(* IEC 61131-3 sources: plc-st-coding-agent/progress/evidence/f14_v10_full_20261113/jobs/codex_minimax-m27 (part 2) *)

(* ---- public-hard-02.candidate_01.st ---- *)
FUNCTION_BLOCK FlexibleProcessingControl
VAR_INPUT
    processLength    : USINT;
    sensor1          : BOOL;
    sensor2          : BOOL;
    sensor3          : BOOL;
    sensor4          : BOOL;
    sensor5          : BOOL;
    station1Start    : BOOL;
    station2Complete : BOOL;
    station3Complete : BOOL;
    station4Complete : BOOL;
    processSequence  : ARRAY[1..8] OF USINT;
END_VAR
VAR_OUTPUT
    conveyorLeft  : BOOL;
    conveyorRight : BOOL;
END_VAR
VAR
    currentState   : UINT := 0;
    currentStation : USINT := 1;
    currentStep    : USINT := 0;
    targetStation  : USINT;
    arrivedAtTarget : BOOL;
    tmpComplete    : BOOL;
END_VAR

(* ENGINEERING_CONTRACT
   State machine with 4 states: IDLE, MOVING, PROCESSING, DONE.
   - PUB001 §3: Start trigger requires sensor1 AND station1Start asserted same scan.
   - PUB002 §3: Conveyor moves to processSequence[currentStep] target station.
   - PUB002 §4: Conveyor stops when target station sensor detects product same scan.
   - PUB003 §5: After arrival, wait for station2Complete/station3Complete/station4Complete.
   - PUB003 §6: Query next sequence element after processing complete same scan.
   - PUB003 §7: Repeat until target is station 5.
   - PUB005 §2: processLength 1..8; processSequence[1..processLength] active.
   - PUB005 §2: Final active entry is station 5; others are stations 2..4.
   - No explicit reset/deactivation required; cycle completes at station 5.
   - No retention of outputs beyond their active state; conveyorLeft/Right only active during MOVING.
   - Direction: targetStation > currentStation → conveyorRight; targetStation < currentStation → conveyorLeft.
   - First movement: from station 1 to processSequence[1].
*)
(* CONTRACT_RULES [] *)

CONST
    STATE_IDLE       := 0;
    STATE_MOVING     := 1;
    STATE_PROCESSING := 2;
    STATE_DONE       := 3;
END_CONST

CASE currentState OF
    STATE_IDLE:
        IF sensor1 AND station1Start THEN
            currentStep := 1;
            currentState := STATE_MOVING;
        END_IF;

    STATE_MOVING:
        targetStation := processSequence[currentStep];

        IF targetStation > currentStation THEN
            conveyorRight := TRUE;
            conveyorLeft := FALSE;
        ELSIF targetStation < currentStation THEN
            conveyorLeft := TRUE;
            conveyorRight := FALSE;
        END_IF;

        arrivedAtTarget :=
            (targetStation = 2 AND sensor2) OR
            (targetStation = 3 AND sensor3) OR
            (targetStation = 4 AND sensor4) OR
            (targetStation = 5 AND sensor5);

        IF arrivedAtTarget THEN
            conveyorLeft := FALSE;
            conveyorRight := FALSE;
            currentStation := targetStation;

            IF targetStation = 5 THEN
                currentState := STATE_DONE;
            ELSE
                currentState := STATE_PROCESSING;
            END_IF;
        END_IF;

    STATE_PROCESSING:
        tmpComplete := FALSE;
        IF currentStation = 2 THEN
            tmpComplete := station2Complete;
        ELSIF currentStation = 3 THEN
            tmpComplete := station3Complete;
        ELSIF currentStation = 4 THEN
            tmpComplete := station4Complete;
        END_IF;

        IF tmpComplete THEN
            currentStep := currentStep + 1;
            currentState := STATE_MOVING;
        END_IF;

    STATE_DONE:

END_CASE;

END_FUNCTION_BLOCK

(* ---- public-hard-02.candidate_02.st ---- *)
FUNCTION_BLOCK FlexibleProcessingControl
VAR_INPUT
    processLength    : USINT;
    sensor1          : BOOL;
    sensor2          : BOOL;
    sensor3          : BOOL;
    sensor4          : BOOL;
    sensor5          : BOOL;
    station1Start    : BOOL;
    station2Complete : BOOL;
    station3Complete : BOOL;
    station4Complete : BOOL;
    processSequence  : ARRAY[1..8] OF USINT;
END_VAR
VAR_OUTPUT
    conveyorLeft  : BOOL;
    conveyorRight : BOOL;
END_VAR
VAR
    currentState   : UINT := 0;
    currentStation : USINT := 1;
    currentStep    : USINT := 0;
    targetStation  : USINT;
    arrivedAtTarget : BOOL;
    tmpComplete    : BOOL;
END_VAR
VAR_CONSTANT
    STATE_IDLE       : UINT := 0;
    STATE_MOVING     : UINT := 1;
    STATE_PROCESSING : UINT := 2;
    STATE_DONE       : UINT := 3;
END_VAR

(* ENGINEERING_CONTRACT
   State machine with 4 states: IDLE, MOVING, PROCESSING, DONE.
   - PUB001 §3: Start trigger requires sensor1 AND station1Start asserted same scan.
   - PUB002 §3: Conveyor moves to processSequence[currentStep] target station.
   - PUB002 §4: Conveyor stops when target station sensor detects product same scan.
   - PUB003 §5: After arrival, wait for station2Complete/station3Complete/station4Complete.
   - PUB003 §6: Query next sequence element after processing complete same scan.
   - PUB003 §7: Repeat until target is station 5.
   - PUB005 §2: processLength 1..8; processSequence[1..processLength] active.
   - PUB005 §2: Final active entry is station 5; others are stations 2..4.
   - No explicit reset/deactivation required; cycle completes at station 5.
   - No retention of outputs beyond their active state; conveyorLeft/Right only active during MOVING.
   - Direction: targetStation > currentStation → conveyorRight; targetStation < currentStation → conveyorLeft.
   - First movement: from station 1 to processSequence[1].
*)
(* CONTRACT_RULES [] *)

CASE currentState OF
    STATE_IDLE:
        IF sensor1 AND station1Start THEN
            currentStep := 1;
            currentState := STATE_MOVING;
        END_IF;

    STATE_MOVING:
        targetStation := processSequence[currentStep];

        IF targetStation > currentStation THEN
            conveyorRight := TRUE;
            conveyorLeft := FALSE;
        ELSIF targetStation < currentStation THEN
            conveyorLeft := TRUE;
            conveyorRight := FALSE;
        END_IF;

        arrivedAtTarget :=
            (targetStation = 2 AND sensor2) OR
            (targetStation = 3 AND sensor3) OR
            (targetStation = 4 AND sensor4) OR
            (targetStation = 5 AND sensor5);

        IF arrivedAtTarget THEN
            conveyorLeft := FALSE;
            conveyorRight := FALSE;
            currentStation := targetStation;

            IF targetStation = 5 THEN
                currentState := STATE_DONE;
            ELSE
                currentState := STATE_PROCESSING;
            END_IF;
        END_IF;

    STATE_PROCESSING:
        tmpComplete := FALSE;
        IF currentStation = 2 THEN
            tmpComplete := station2Complete;
        ELSIF currentStation = 3 THEN
            tmpComplete := station3Complete;
        ELSIF currentStation = 4 THEN
            tmpComplete := station4Complete;
        END_IF;

        IF tmpComplete THEN
            currentStep := currentStep + 1;
            currentState := STATE_MOVING;
        END_IF;

    STATE_DONE:

END_CASE;

END_FUNCTION_BLOCK

(* ---- public-hard-02.candidate_03.st ---- *)
FUNCTION_BLOCK FlexibleProcessingControl
VAR_INPUT
    processLength    : USINT;
    sensor1          : BOOL;
    sensor2          : BOOL;
    sensor3          : BOOL;
    sensor4          : BOOL;
    sensor5          : BOOL;
    station1Start    : BOOL;
    station2Complete : BOOL;
    station3Complete : BOOL;
    station4Complete : BOOL;
    processSequence  : ARRAY[1..8] OF USINT;
END_VAR
VAR_OUTPUT
    conveyorLeft  : BOOL;
    conveyorRight : BOOL;
END_VAR
VAR
    currentState   : UINT := 0;
    currentStation : USINT := 1;
    currentStep    : USINT := 0;
    targetStation  : USINT;
    arrivedAtTarget : BOOL;
    tmpComplete    : BOOL;
END_VAR

(* ENGINEERING_CONTRACT
   State machine with 4 states: IDLE, MOVING, PROCESSING, DONE.
   - PUB001 §3: Start trigger requires sensor1 AND station1Start asserted same scan.
   - PUB002 §3: Conveyor moves to processSequence[currentStep] target station.
   - PUB002 §4: Conveyor stops when target station sensor detects product same scan.
   - PUB003 §5: After arrival, wait for station2Complete/station3Complete/station4Complete.
   - PUB003 §6: Query next sequence element after processing complete same scan.
   - PUB003 §7: Repeat until target is station 5.
   - PUB005 §2: processLength 1..8; processSequence[1..processLength] active.
   - PUB005 §2: Final active entry is station 5; others are stations 2..4.
   - No explicit reset/deactivation required; cycle completes at station 5.
   - No retention of outputs beyond their active state; conveyorLeft/Right only active during MOVING.
   - Direction: targetStation > currentStation → conveyorRight; targetStation < currentStation → conveyorLeft.
   - First movement: from station 1 to processSequence[1].
*)
(* CONTRACT_RULES [] *)

CASE currentState OF
    0: (* IDLE *)
        IF sensor1 AND station1Start THEN
            currentStep := 1;
            currentState := 1;
        END_IF;

    1: (* MOVING *)
        targetStation := processSequence[currentStep];

        IF targetStation > currentStation THEN
            conveyorRight := TRUE;
            conveyorLeft := FALSE;
        ELSIF targetStation < currentStation THEN
            conveyorLeft := TRUE;
            conveyorRight := FALSE;
        END_IF;

        arrivedAtTarget :=
            (targetStation = 2 AND sensor2) OR
            (targetStation = 3 AND sensor3) OR
            (targetStation = 4 AND sensor4) OR
            (targetStation = 5 AND sensor5);

        IF arrivedAtTarget THEN
            conveyorLeft := FALSE;
            conveyorRight := FALSE;
            currentStation := targetStation;

            IF targetStation = 5 THEN
                currentState := 3;
            ELSE
                currentState := 2;
            END_IF;
        END_IF;

    2: (* PROCESSING *)
        tmpComplete := FALSE;
        IF currentStation = 2 THEN
            tmpComplete := station2Complete;
        ELSIF currentStation = 3 THEN
            tmpComplete := station3Complete;
        ELSIF currentStation = 4 THEN
            tmpComplete := station4Complete;
        END_IF;

        IF tmpComplete THEN
            currentStep := currentStep + 1;
            currentState := 1;
        END_IF;

    3: (* DONE *)

END_CASE;

END_FUNCTION_BLOCK

(* ---- public-hard-02.candidate_04.st ---- *)
FUNCTION_BLOCK FlexibleProcessingControl
VAR_INPUT
    processLength    : USINT;
    sensor1          : BOOL;
    sensor2          : BOOL;
    sensor3          : BOOL;
    sensor4          : BOOL;
    sensor5          : BOOL;
    station1Start    : BOOL;
    station2Complete : BOOL;
    station3Complete : BOOL;
    station4Complete : BOOL;
    processSequence  : ARRAY[1..8] OF USINT;
END_VAR
VAR_OUTPUT
    conveyorLeft  : BOOL;
    conveyorRight : BOOL;
END_VAR
VAR
    currentState   : UINT := 0;
    currentStation : USINT := 1;
    currentStep    : USINT := 0;
    tmp_target     : USINT;
    tmp_arrived    : BOOL;
    tmp_complete   : BOOL;
END_VAR

(* ENGINEERING_CONTRACT
   State machine: IDLE(0), MOVING(1), PROCESSING(2), DONE(3).
   - PUB001 §1: 5 workstations, 1#=load, 2-4#=process, 5#=output.
   - PUB005 §3: Start requires sensor1 AND station1Start same scan.
   - PUB005 §3: Query processSequence[1], start conveyor to target.
   - PUB005 §4: Stop conveyor when target station sensor detects product.
   - PUB005 §5: Wait for station2Complete/station3Complete/station4Complete.
   - PUB005 §6: After completion, query next processSequence element.
   - PUB005 §7: Repeat until target is station 5.
   - PUB005 §2: processLength 1..8; final entry=5, others=2..4.
   - No explicit reset; cycle completes at station 5.
   - conveyorLeft/Right active only during MOVING to target.
   - Direction: target > current → Right; target < current → Left.
   - currentStation tracks physical position; updates on arrival only.
*)
(* CONTRACT_RULES [] *)

CASE currentState OF
    0: (* IDLE *)
        IF sensor1 AND station1Start THEN
            currentStep := 1;
            currentState := 1;
        END_IF;

    1: (* MOVING *)
        tmp_target := processSequence[currentStep];

        IF tmp_target > currentStation THEN
            conveyorRight := TRUE;
            conveyorLeft := FALSE;
        ELSIF tmp_target < currentStation THEN
            conveyorLeft := TRUE;
            conveyorRight := FALSE;
        ELSE
            conveyorRight := FALSE;
            conveyorLeft := FALSE;
        END_IF;

        tmp_arrived :=
            (tmp_target = 2 AND sensor2) OR
            (tmp_target = 3 AND sensor3) OR
            (tmp_target = 4 AND sensor4) OR
            (tmp_target = 5 AND sensor5);

        IF tmp_arrived THEN
            conveyorLeft := FALSE;
            conveyorRight := FALSE;
            currentStation := tmp_target;

            IF tmp_target = 5 THEN
                currentState := 3;
            ELSE
                currentState := 2;
            END_IF;
        END_IF;

    2: (* PROCESSING *)
        tmp_complete := FALSE;
        IF currentStation = 2 THEN
            tmp_complete := station2Complete;
        ELSIF currentStation = 3 THEN
            tmp_complete := station3Complete;
        ELSIF currentStation = 4 THEN
            tmp_complete := station4Complete;
        END_IF;

        IF tmp_complete THEN
            currentStep := currentStep + 1;
            currentState := 1;
        END_IF;

    3: (* DONE *)

END_CASE;

END_FUNCTION_BLOCK

(* ---- public-hard-02.raw_candidate_01.st ---- *)
FUNCTION_BLOCK FlexibleProcessingControl
VAR_INPUT
    processLength    : USINT;
    sensor1          : BOOL;
    sensor2          : BOOL;
    sensor3          : BOOL;
    sensor4          : BOOL;
    sensor5          : BOOL;
    station1Start    : BOOL;
    station2Complete : BOOL;
    station3Complete : BOOL;
    station4Complete : BOOL;
    processSequence  : ARRAY[1..8] OF USINT;
END_VAR
VAR_OUTPUT
    conveyorLeft  : BOOL;
    conveyorRight : BOOL;
END_VAR
VAR
    currentState   : UINT := 0;
    currentStation : USINT := 1;
    currentStep    : USINT := 0;
    targetStation  : USINT;
    arrivedAtTarget : BOOL;
    tmpComplete    : BOOL;
END_VAR

(* ENGINEERING_CONTRACT
   State machine with 4 states: IDLE, MOVING, PROCESSING, DONE.
   - PUB001 §3: Start trigger requires sensor1 AND station1Start asserted same scan.
   - PUB002 §3: Conveyor moves to processSequence[currentStep] target station.
   - PUB002 §4: Conveyor stops when target station sensor detects product same scan.
   - PUB003 §5: After arrival, wait for station2Complete/station3Complete/station4Complete.
   - PUB003 §6: Query next sequence element after processing complete same scan.
   - PUB003 §7: Repeat until target is station 5.
   - PUB005 §2: processLength 1..8; processSequence[1..processLength] active.
   - PUB005 §2: Final active entry is station 5; others are stations 2..4.
   - No explicit reset/deactivation required; cycle completes at station 5.
   - No retention of outputs beyond their active state; conveyorLeft/Right only active during MOVING.
   - Direction: targetStation > currentStation → conveyorRight; targetStation < currentStation → conveyorLeft.
   - First movement: from station 1 to processSequence[1].
*)
(* CONTRACT_RULES [] *)

CONST
    STATE_IDLE       := 0;
    STATE_MOVING     := 1;
    STATE_PROCESSING := 2;
    STATE_DONE       := 3;
END_CONST

CASE currentState OF
    STATE_IDLE:
        IF sensor1 AND station1Start THEN
            currentStep := 1;
            currentState := STATE_MOVING;
        END_IF;

    STATE_MOVING:
        targetStation := processSequence[currentStep];

        IF targetStation > currentStation THEN
            conveyorRight := TRUE;
            conveyorLeft := FALSE;
        ELSIF targetStation < currentStation THEN
            conveyorLeft := TRUE;
            conveyorRight := FALSE;
        END_IF;

        arrivedAtTarget :=
            (targetStation = 2 AND sensor2) OR
            (targetStation = 3 AND sensor3) OR
            (targetStation = 4 AND sensor4) OR
            (targetStation = 5 AND sensor5);

        IF arrivedAtTarget THEN
            conveyorLeft := FALSE;
            conveyorRight := FALSE;
            currentStation := targetStation;

            IF targetStation = 5 THEN
                currentState := STATE_DONE;
            ELSE
                currentState := STATE_PROCESSING;
            END_IF;
        END_IF;

    STATE_PROCESSING:
        tmpComplete := FALSE;
        IF currentStation = 2 THEN
            tmpComplete := station2Complete;
        ELSIF currentStation = 3 THEN
            tmpComplete := station3Complete;
        ELSIF currentStation = 4 THEN
            tmpComplete := station4Complete;
        END_IF;

        IF tmpComplete THEN
            currentStep := currentStep + 1;
            currentState := STATE_MOVING;
        END_IF;

    STATE_DONE:

END_CASE;

END_FUNCTION_BLOCK

(* ---- public-hard-02.raw_candidate_02.st ---- *)
FUNCTION_BLOCK FlexibleProcessingControl
VAR_INPUT
    processLength    : USINT;
    sensor1          : BOOL;
    sensor2          : BOOL;
    sensor3          : BOOL;
    sensor4          : BOOL;
    sensor5          : BOOL;
    station1Start    : BOOL;
    station2Complete : BOOL;
    station3Complete : BOOL;
    station4Complete : BOOL;
    processSequence  : ARRAY[1..8] OF USINT;
END_VAR
VAR_OUTPUT
    conveyorLeft  : BOOL;
    conveyorRight : BOOL;
END_VAR
VAR
    currentState   : UINT := 0;
    currentStation : USINT := 1;
    currentStep    : USINT := 0;
    targetStation  : USINT;
    arrivedAtTarget : BOOL;
    tmpComplete    : BOOL;
END_VAR
VAR_CONSTANT
    STATE_IDLE       : UINT := 0;
    STATE_MOVING     : UINT := 1;
    STATE_PROCESSING : UINT := 2;
    STATE_DONE       : UINT := 3;
END_VAR

(* ENGINEERING_CONTRACT
   State machine with 4 states: IDLE, MOVING, PROCESSING, DONE.
   - PUB001 §3: Start trigger requires sensor1 AND station1Start asserted same scan.
   - PUB002 §3: Conveyor moves to processSequence[currentStep] target station.
   - PUB002 §4: Conveyor stops when target station sensor detects product same scan.
   - PUB003 §5: After arrival, wait for station2Complete/station3Complete/station4Complete.
   - PUB003 §6: Query next sequence element after processing complete same scan.
   - PUB003 §7: Repeat until target is station 5.
   - PUB005 §2: processLength 1..8; processSequence[1..processLength] active.
   - PUB005 §2: Final active entry is station 5; others are stations 2..4.
   - No explicit reset/deactivation required; cycle completes at station 5.
   - No retention of outputs beyond their active state; conveyorLeft/Right only active during MOVING.
   - Direction: targetStation > currentStation → conveyorRight; targetStation < currentStation → conveyorLeft.
   - First movement: from station 1 to processSequence[1].
*)
(* CONTRACT_RULES [] *)

CASE currentState OF
    STATE_IDLE:
        IF sensor1 AND station1Start THEN
            currentStep := 1;
            currentState := STATE_MOVING;
        END_IF;

    STATE_MOVING:
        targetStation := processSequence[currentStep];

        IF targetStation > currentStation THEN
            conveyorRight := TRUE;
            conveyorLeft := FALSE;
        ELSIF targetStation < currentStation THEN
            conveyorLeft := TRUE;
            conveyorRight := FALSE;
        END_IF;

        arrivedAtTarget :=
            (targetStation = 2 AND sensor2) OR
            (targetStation = 3 AND sensor3) OR
            (targetStation = 4 AND sensor4) OR
            (targetStation = 5 AND sensor5);

        IF arrivedAtTarget THEN
            conveyorLeft := FALSE;
            conveyorRight := FALSE;
            currentStation := targetStation;

            IF targetStation = 5 THEN
                currentState := STATE_DONE;
            ELSE
                currentState := STATE_PROCESSING;
            END_IF;
        END_IF;

    STATE_PROCESSING:
        tmpComplete := FALSE;
        IF currentStation = 2 THEN
            tmpComplete := station2Complete;
        ELSIF currentStation = 3 THEN
            tmpComplete := station3Complete;
        ELSIF currentStation = 4 THEN
            tmpComplete := station4Complete;
        END_IF;

        IF tmpComplete THEN
            currentStep := currentStep + 1;
            currentState := STATE_MOVING;
        END_IF;

    STATE_DONE:

END_CASE;

END_FUNCTION_BLOCK

(* ---- public-hard-02.raw_candidate_03.st ---- *)
FUNCTION_BLOCK FlexibleProcessingControl
VAR_INPUT
    processLength    : USINT;
    sensor1          : BOOL;
    sensor2          : BOOL;
    sensor3          : BOOL;
    sensor4          : BOOL;
    sensor5          : BOOL;
    station1Start    : BOOL;
    station2Complete : BOOL;
    station3Complete : BOOL;
    station4Complete : BOOL;
    processSequence  : ARRAY[1..8] OF USINT;
END_VAR
VAR_OUTPUT
    conveyorLeft  : BOOL;
    conveyorRight : BOOL;
END_VAR
VAR
    currentState   : UINT := 0;
    currentStation : USINT := 1;
    currentStep    : USINT := 0;
    targetStation  : USINT;
    arrivedAtTarget : BOOL;
    tmpComplete    : BOOL;
END_VAR

(* ENGINEERING_CONTRACT
   State machine with 4 states: IDLE, MOVING, PROCESSING, DONE.
   - PUB001 §3: Start trigger requires sensor1 AND station1Start asserted same scan.
   - PUB002 §3: Conveyor moves to processSequence[currentStep] target station.
   - PUB002 §4: Conveyor stops when target station sensor detects product same scan.
   - PUB003 §5: After arrival, wait for station2Complete/station3Complete/station4Complete.
   - PUB003 §6: Query next sequence element after processing complete same scan.
   - PUB003 §7: Repeat until target is station 5.
   - PUB005 §2: processLength 1..8; processSequence[1..processLength] active.
   - PUB005 §2: Final active entry is station 5; others are stations 2..4.
   - No explicit reset/deactivation required; cycle completes at station 5.
   - No retention of outputs beyond their active state; conveyorLeft/Right only active during MOVING.
   - Direction: targetStation > currentStation → conveyorRight; targetStation < currentStation → conveyorLeft.
   - First movement: from station 1 to processSequence[1].
*)
(* CONTRACT_RULES [] *)

CASE currentState OF
    0: (* IDLE *)
        IF sensor1 AND station1Start THEN
            currentStep := 1;
            currentState := 1;
        END_IF;

    1: (* MOVING *)
        targetStation := processSequence[currentStep];

        IF targetStation > currentStation THEN
            conveyorRight := TRUE;
            conveyorLeft := FALSE;
        ELSIF targetStation < currentStation THEN
            conveyorLeft := TRUE;
            conveyorRight := FALSE;
        END_IF;

        arrivedAtTarget :=
            (targetStation = 2 AND sensor2) OR
            (targetStation = 3 AND sensor3) OR
            (targetStation = 4 AND sensor4) OR
            (targetStation = 5 AND sensor5);

        IF arrivedAtTarget THEN
            conveyorLeft := FALSE;
            conveyorRight := FALSE;
            currentStation := targetStation;

            IF targetStation = 5 THEN
                currentState := 3;
            ELSE
                currentState := 2;
            END_IF;
        END_IF;

    2: (* PROCESSING *)
        tmpComplete := FALSE;
        IF currentStation = 2 THEN
            tmpComplete := station2Complete;
        ELSIF currentStation = 3 THEN
            tmpComplete := station3Complete;
        ELSIF currentStation = 4 THEN
            tmpComplete := station4Complete;
        END_IF;

        IF tmpComplete THEN
            currentStep := currentStep + 1;
            currentState := 1;
        END_IF;

    3: (* DONE *)

END_CASE;

END_FUNCTION_BLOCK

(* ---- public-hard-02.raw_candidate_04.st ---- *)
FUNCTION_BLOCK FlexibleProcessingControl
VAR_INPUT
    processLength    : USINT;
    sensor1          : BOOL;
    sensor2          : BOOL;
    sensor3          : BOOL;
    sensor4          : BOOL;
    sensor5          : BOOL;
    station1Start    : BOOL;
    station2Complete : BOOL;
    station3Complete : BOOL;
    station4Complete : BOOL;
    processSequence  : ARRAY[1..8] OF USINT;
END_VAR
VAR_OUTPUT
    conveyorLeft  : BOOL;
    conveyorRight : BOOL;
END_VAR
VAR
    currentState   : UINT := 0;
    currentStation : USINT := 1;
    currentStep    : USINT := 0;
    tmp_target     : USINT;
    tmp_arrived    : BOOL;
    tmp_complete   : BOOL;
END_VAR

(* ENGINEERING_CONTRACT
   State machine: IDLE(0), MOVING(1), PROCESSING(2), DONE(3).
   - PUB001 §1: 5 workstations, 1#=load, 2-4#=process, 5#=output.
   - PUB005 §3: Start requires sensor1 AND station1Start same scan.
   - PUB005 §3: Query processSequence[1], start conveyor to target.
   - PUB005 §4: Stop conveyor when target station sensor detects product.
   - PUB005 §5: Wait for station2Complete/station3Complete/station4Complete.
   - PUB005 §6: After completion, query next processSequence element.
   - PUB005 §7: Repeat until target is station 5.
   - PUB005 §2: processLength 1..8; final entry=5, others=2..4.
   - No explicit reset; cycle completes at station 5.
   - conveyorLeft/Right active only during MOVING to target.
   - Direction: target > current → Right; target < current → Left.
   - currentStation tracks physical position; updates on arrival only.
*)
(* CONTRACT_RULES [] *)

CASE currentState OF
    0: (* IDLE *)
        IF sensor1 AND station1Start THEN
            currentStep := 1;
            currentState := 1;
        END_IF;

    1: (* MOVING *)
        tmp_target := processSequence[currentStep];

        IF tmp_target > currentStation THEN
            conveyorRight := TRUE;
            conveyorLeft := FALSE;
        ELSIF tmp_target < currentStation THEN
            conveyorLeft := TRUE;
            conveyorRight := FALSE;
        ELSE
            conveyorRight := FALSE;
            conveyorLeft := FALSE;
        END_IF;

        tmp_arrived :=
            (tmp_target = 2 AND sensor2) OR
            (tmp_target = 3 AND sensor3) OR
            (tmp_target = 4 AND sensor4) OR
            (tmp_target = 5 AND sensor5);

        IF tmp_arrived THEN
            conveyorLeft := FALSE;
            conveyorRight := FALSE;
            currentStation := tmp_target;

            IF tmp_target = 5 THEN
                currentState := 3;
            ELSE
                currentState := 2;
            END_IF;
        END_IF;

    2: (* PROCESSING *)
        tmp_complete := FALSE;
        IF currentStation = 2 THEN
            tmp_complete := station2Complete;
        ELSIF currentStation = 3 THEN
            tmp_complete := station3Complete;
        ELSIF currentStation = 4 THEN
            tmp_complete := station4Complete;
        END_IF;

        IF tmp_complete THEN
            currentStep := currentStep + 1;
            currentState := 1;
        END_IF;

    3: (* DONE *)

END_CASE;

END_FUNCTION_BLOCK

(* ---- public-hard-03.candidate_01.st ---- *)
{+
Engineer: Claude
Date: 2026-11-13
Purpose: Recipe Management System per task specification
-}
FUNCTION_BLOCK FB_RecipeManager
VAR_INPUT
    addRecipe    : BOOL;
    deleteRecipe : BOOL;
    modifyRecipe : BOOL;
    queryRecipe  : BOOL;
    recipeIn     : ST_Recipe;
END_VAR
VAR_OUTPUT
    recipeAdded       : BOOL := FALSE;
    recipeDeleted     : BOOL := FALSE;
    recipeModified    : BOOL := FALSE;
    error             : BOOL := FALSE;
    status            : WORD := 16#0000;
    recipeQueryResult : ST_Recipe;
END_VAR
VAR_IN_OUT
    recipe : ARRAY[1..10] OF ST_Recipe;
END_VAR
VAR
    tmp_index     : INT;
    tmp_found     : BOOL;
    tmp_emptySlot : INT;
    tmp_hasEmpty  : BOOL;
END_VAR

(*
ENGINEERING_CONTRACT
====================
Operation Execution (same-scan, sequential priority order):
1. queryRecipe  → PUB001, PUB002, PUB008
2. addRecipe    → PUB002, PUB003, PUB009
3. deleteRecipe → PUB002, PUB004, PUB010
4. modifyRecipe → PUB002, PUB005, PUB011

Outputs - Activation/Retention/Reset:
- recipeAdded/recipeDeleted/recipeModified: pulse TRUE on success for current scan only (no retention)
- error: TRUE when any error occurs; no explicit reset (overwritten next scan)
- status: 16#0000 no-error, or error code 16#8001-16#8005 per PUB002

Error Codes (PUB002):
- 16#8001: queryRecipe - recipeID not found
- 16#8002: addRecipe   - recipeID already exists (duplicate)
- 16#8003: addRecipe   - no empty slot (database full)
- 16#8004: deleteRecipe - recipeID not found
- 16#8005: modifyRecipe - recipeID not found

Database Semantics (PUB006, PUB007):
- Array index range: [1..10], fixed
- Empty slot: recipeID = 0
- Add stores at smallest index empty slot (lowest array index)
- Delete sets recipeID to 0 (marks slot empty)
- Duplicate recipeID prohibited

Boundary Checks:
- recipeID comparisons use exact equality
- No wraparound or saturation logic
*)

(* CONTRACT_RULES [] *)

recipeAdded    := FALSE;
recipeDeleted  := FALSE;
recipeModified := FALSE;
error          := FALSE;
status         := 16#0000;

IF queryRecipe THEN
    tmp_found  := FALSE;
    tmp_index  := 1;
    FOR tmp_index := 1 TO 10 DO
        IF recipe[tmp_index].recipeID = recipeIn.recipeID THEN
            tmp_found := TRUE;
            EXIT;
        END_IF
    END_FOR;

    IF tmp_found THEN
        recipeQueryResult := recipe[tmp_index];
    ELSE
        error  := TRUE;
        status := 16#8001;
    END_IF;
END_IF;

IF addRecipe THEN
    tmp_found     := FALSE;
    tmp_hasEmpty  := FALSE;
    tmp_emptySlot := 0;

    FOR tmp_index := 1 TO 10 DO
        IF recipe[tmp_index].recipeID = recipeIn.recipeID THEN
            tmp_found := TRUE;
            EXIT;
        END_IF;
        IF recipe[tmp_index].recipeID = 0 AND NOT tmp_hasEmpty THEN
            tmp_hasEmpty  := TRUE;
            tmp_emptySlot := tmp_index;
        END_IF;
    END_FOR;

    IF tmp_found THEN
        error  := TRUE;
        status := 16#8002;
    ELSIF NOT tmp_hasEmpty THEN
        error  := TRUE;
        status := 16#8003;
    ELSE
        recipe[tmp_emptySlot] := recipeIn;
        recipeAdded           := TRUE;
    END_IF;
END_IF;

IF deleteRecipe THEN
    tmp_found := FALSE;
    tmp_index := 1;

    FOR tmp_index := 1 TO 10 DO
        IF recipe[tmp_index].recipeID = recipeIn.recipeID THEN
            tmp_found := TRUE;
            EXIT;
        END_IF;
    END_FOR;

    IF tmp_found THEN
        recipe[tmp_index].recipeID := 0;
        recipeDeleted              := TRUE;
    ELSE
        error  := TRUE;
        status := 16#8004;
    END_IF;
END_IF;

IF modifyRecipe THEN
    tmp_found := FALSE;
    tmp_index := 1;

    FOR tmp_index := 1 TO 10 DO
        IF recipe[tmp_index].recipeID = recipeIn.recipeID THEN
            tmp_found := TRUE;
            EXIT;
        END_IF;
    END_FOR;

    IF tmp_found THEN
        recipe[tmp_index] := recipeIn;
        recipeModified    := TRUE;
    ELSE
        error  := TRUE;
        status := 16#8005;
    END_IF;
END_IF;

END_FUNCTION_BLOCK

(* ---- public-hard-03.candidate_02.st ---- *)
{+
FUNCTION_BLOCK FB_RecipeManager
VAR_INPUT
    addRecipe    : BOOL;
    deleteRecipe : BOOL;
    modifyRecipe : BOOL;
    queryRecipe  : BOOL;
    recipeIn     : ST_Recipe;
END_VAR
VAR_OUTPUT
    recipeAdded       : BOOL := FALSE;
    recipeDeleted     : BOOL := FALSE;
    recipeModified    : BOOL := FALSE;
    error             : BOOL := FALSE;
    status            : WORD := 16#0000;
    recipeQueryResult : ST_Recipe;
END_VAR
VAR_IN_OUT
    recipe : ARRAY[1..10] OF ST_Recipe;
END_VAR
VAR
    tmp_index     : INT;
    tmp_found     : BOOL;
    tmp_emptySlot : INT;
    tmp_hasEmpty  : BOOL;
END_VAR

(* ENGINEERING_CONTRACT
   ====================
   Operation Execution (same-scan, sequential priority):
   1. queryRecipe  → PUB008
   2. addRecipe    → PUB009
   3. deleteRecipe → PUB010
   4. modifyRecipe → PUB011

   Outputs - Activation/Retention/Reset:
   - recipeAdded/recipeDeleted/recipeModified: pulse TRUE on success for current scan only
   - error: TRUE when any error occurs; no explicit reset (overwritten next scan)
   - status: 16#0000 no-error, or error code 16#8001-16#8005 per PUB002

   Error Codes (PUB002):
   - 16#8001: queryRecipe - recipeID not found
   - 16#8002: addRecipe   - recipeID already exists (duplicate)
   - 16#8003: addRecipe   - no empty slot (database full)
   - 16#8004: deleteRecipe - recipeID not found
   - 16#8005: modifyRecipe - recipeID not found

   Database Semantics (PUB006, PUB007):
   - Array index range: [1..10], fixed
   - Empty slot: recipeID = 0
   - Add stores at smallest index empty slot
   - Delete sets recipeID to 0 (marks slot empty)
   - Duplicate recipeID prohibited
*)

(* CONTRACT_RULES [] *)

recipeAdded    := FALSE;
recipeDeleted  := FALSE;
recipeModified := FALSE;
error          := FALSE;
status         := 16#0000;

IF queryRecipe THEN
    tmp_found := FALSE;
    tmp_index := 1;
    WHILE tmp_index <= 10 AND NOT tmp_found DO
        IF recipe[tmp_index].recipeID = recipeIn.recipeID THEN
            tmp_found := TRUE;
        ELSE
            tmp_index := tmp_index + 1;
        END_IF;
    END_WHILE;

    IF tmp_found THEN
        recipeQueryResult := recipe[tmp_index];
    ELSE
        error  := TRUE;
        status := 16#8001;
    END_IF;
END_IF;

IF addRecipe THEN
    tmp_found     := FALSE;
    tmp_hasEmpty  := FALSE;
    tmp_emptySlot := 0;
    tmp_index     := 1;

    WHILE tmp_index <= 10 DO
        IF recipe[tmp_index].recipeID = recipeIn.recipeID THEN
            tmp_found := TRUE;
            tmp_index := 11;
        ELSE
            IF recipe[tmp_index].recipeID = 0 AND NOT tmp_hasEmpty THEN
                tmp_hasEmpty  := TRUE;
                tmp_emptySlot := tmp_index;
            END_IF;
            tmp_index := tmp_index + 1;
        END_IF;
    END_WHILE;

    IF tmp_found THEN
        error  := TRUE;
        status := 16#8002;
    ELSIF NOT tmp_hasEmpty THEN
        error  := TRUE;
        status := 16#8003;
    ELSE
        recipe[tmp_emptySlot] := recipeIn;
        recipeAdded           := TRUE;
    END_IF;
END_IF;

IF deleteRecipe THEN
    tmp_found := FALSE;
    tmp_index := 1;

    WHILE tmp_index <= 10 AND NOT tmp_found DO
        IF recipe[tmp_index].recipeID = recipeIn.recipeID THEN
            tmp_found := TRUE;
        ELSE
            tmp_index := tmp_index + 1;
        END_IF;
    END_WHILE;

    IF tmp_found THEN
        recipe[tmp_index].recipeID := 0;
        recipeDeleted              := TRUE;
    ELSE
        error  := TRUE;
        status := 16#8004;
    END_IF;
END_IF;

IF modifyRecipe THEN
    tmp_found := FALSE;
    tmp_index := 1;

    WHILE tmp_index <= 10 AND NOT tmp_found DO
        IF recipe[tmp_index].recipeID = recipeIn.recipeID THEN
            tmp_found := TRUE;
        ELSE
            tmp_index := tmp_index + 1;
        END_IF;
    END_WHILE;

    IF tmp_found THEN
        recipe[tmp_index] := recipeIn;
        recipeModified    := TRUE;
    ELSE
        error  := TRUE;
        status := 16#8005;
    END_IF;
END_IF;

END_FUNCTION_BLOCK
}

(* ---- public-hard-03.candidate_03.st ---- *)
TYPE ST_Recipe :
STRUCT
    recipeID              : INT;
    ingredientType        : INT;
    ingredientRatio       : REAL;
    productionTemperature : REAL;
END_STRUCT
END_TYPE;

FUNCTION_BLOCK FB_RecipeManager
VAR_INPUT
    addRecipe    : BOOL;
    deleteRecipe : BOOL;
    modifyRecipe : BOOL;
    queryRecipe  : BOOL;
    recipeIn     : ST_Recipe;
END_VAR
VAR_OUTPUT
    recipeAdded       : BOOL := FALSE;
    recipeDeleted     : BOOL := FALSE;
    recipeModified    : BOOL := FALSE;
    error             : BOOL := FALSE;
    status            : WORD := 16#0000;
    recipeQueryResult : ST_Recipe;
END_VAR
VAR_IN_OUT
    recipe : ARRAY[1..10] OF ST_Recipe;
END_VAR
VAR
    tmp_index     : INT;
    tmp_found     : BOOL;
    tmp_emptySlot : INT;
    tmp_hasEmpty  : BOOL;
END_VAR

(*
ENGINEERING_CONTRACT
====================
Operation Execution (same-scan, sequential priority order):
1. queryRecipe  -> PUB001, PUB002, PUB008
2. addRecipe    -> PUB002, PUB003, PUB009
3. deleteRecipe -> PUB002, PUB004, PUB010
4. modifyRecipe -> PUB002, PUB005, PUB011

Outputs - Activation/Retention/Reset:
- recipeAdded/recipeDeleted/recipeModified: pulse TRUE on success for current scan only (no retention)
- error: TRUE when any error occurs; no explicit reset (overwritten next scan)
- status: 16#0000 no-error, or error code 16#8001-16#8005 per PUB002

Error Codes (PUB002):
- 16#8001: queryRecipe - recipeID not found
- 16#8002: addRecipe   - recipeID already exists (duplicate)
- 16#8003: addRecipe   - no empty slot (database full)
- 16#8004: deleteRecipe - recipeID not found
- 16#8005: modifyRecipe - recipeID not found

Database Semantics (PUB006, PUB007):
- Array index range: [1..10], fixed
- Empty slot: recipeID = 0
- Add stores at smallest index empty slot (lowest array index)
- Delete sets recipeID to 0 (marks slot empty)
- Duplicate recipeID prohibited

Boundary Checks:
- recipeID comparisons use exact equality
- No wraparound or saturation logic
*)

(* CONTRACT_RULES [] *)

recipeAdded    := FALSE;
recipeDeleted  := FALSE;
recipeModified := FALSE;
error          := FALSE;
status         := 16#0000;

IF queryRecipe THEN
    tmp_found := FALSE;

    FOR tmp_index := 1 TO 10 DO
        IF recipe[tmp_index].recipeID = recipeIn.recipeID THEN
            tmp_found := TRUE;
            EXIT;
        END_IF;
    END_FOR;

    IF tmp_found THEN
        recipeQueryResult := recipe[tmp_index];
    ELSE
        error  := TRUE;
        status := 16#8001;
    END_IF;
END_IF;

IF addRecipe THEN
    tmp_found     := FALSE;
    tmp_hasEmpty  := FALSE;
    tmp_emptySlot := 0;

    FOR tmp_index := 1 TO 10 DO
        IF recipe[tmp_index].recipeID = recipeIn.recipeID THEN
            tmp_found := TRUE;
            EXIT;
        END_IF;
        IF recipe[tmp_index].recipeID = 0 AND NOT tmp_hasEmpty THEN
            tmp_hasEmpty  := TRUE;
            tmp_emptySlot := tmp_index;
        END_IF;
    END_FOR;

    IF tmp_found THEN
        error  := TRUE;
        status := 16#8002;
    ELSIF NOT tmp_hasEmpty THEN
        error  := TRUE;
        status := 16#8003;
    ELSE
        recipe[tmp_emptySlot] := recipeIn;
        recipeAdded           := TRUE;
    END_IF;
END_IF;

IF deleteRecipe THEN
    tmp_found := FALSE;

    FOR tmp_index := 1 TO 10 DO
        IF recipe[tmp_index].recipeID = recipeIn.recipeID THEN
            tmp_found := TRUE;
            EXIT;
        END_IF;
    END_FOR;

    IF tmp_found THEN
        recipe[tmp_index].recipeID := 0;
        recipeDeleted              := TRUE;
    ELSE
        error  := TRUE;
        status := 16#8004;
    END_IF;
END_IF;

IF modifyRecipe THEN
    tmp_found := FALSE;

    FOR tmp_index := 1 TO 10 DO
        IF recipe[tmp_index].recipeID = recipeIn.recipeID THEN
            tmp_found := TRUE;
            EXIT;
        END_IF;
    END_FOR;

    IF tmp_found THEN
        recipe[tmp_index] := recipeIn;
        recipeModified    := TRUE;
    ELSE
        error  := TRUE;
        status := 16#8005;
    END_IF;
END_IF;

END_FUNCTION_BLOCK

(* ---- public-hard-03.candidate_04.st ---- *)
TYPE ST_Recipe :
STRUCT
    recipeID              : INT;
    ingredientType        : INT;
    ingredientRatio       : REAL;
    productionTemperature : REAL;
END_STRUCT
END_TYPE;

FUNCTION_BLOCK FB_RecipeManager
VAR_INPUT
    addRecipe    : BOOL;
    deleteRecipe : BOOL;
    modifyRecipe : BOOL;
    queryRecipe  : BOOL;
    recipeIn     : ST_Recipe;
END_VAR
VAR_OUTPUT
    recipeAdded       : BOOL := FALSE;
    recipeDeleted     : BOOL := FALSE;
    recipeModified    : BOOL := FALSE;
    error             : BOOL := FALSE;
    status            : WORD := 16#0000;
    recipeQueryResult : ST_Recipe;
END_VAR
VAR_IN_OUT
    recipe : ARRAY[1..10] OF ST_Recipe;
END_VAR
VAR
    local_index         : INT;
    local_found         : BOOL;
    local_emptySlot     : INT;
    local_hasEmpty      : BOOL;
    local_opExecuted    : BOOL;
END_VAR

(*
ENGINEERING_CONTRACT
====================
Operation Execution (same-scan, sequential priority order):
1. queryRecipe  -> PUB001, PUB002, PUB008
2. addRecipe    -> PUB002, PUB003, PUB009
3. deleteRecipe -> PUB002, PUB004, PUB010
4. modifyRecipe -> PUB002, PUB005, PUB011

Outputs - Activation/Retention/Reset:
- recipeAdded/recipeDeleted/recipeModified: pulse TRUE on success for current scan only (no retention)
- error: TRUE when any error occurs; retained across calls until next operation runs
- status: 16#0000 no-error, or error code 16#8001-16#8005 per PUB002; retained across calls

Error Codes (PUB002):
- 16#8001: queryRecipe  - recipeID not found
- 16#8002: addRecipe    - recipeID already exists (duplicate)
- 16#8003: addRecipe    - no empty slot (database full)
- 16#8004: deleteRecipe - recipeID not found
- 16#8005: modifyRecipe - recipeID not found

Database Semantics (PUB006, PUB007):
- Array index range: [1..10], fixed
- Empty slot: recipeID = 0
- Add stores at smallest index empty slot (lowest array index)
- Delete sets recipeID to 0 (marks slot empty)
- Duplicate recipeID prohibited

Boundary Checks:
- recipeID comparisons use exact equality
- No wraparound or saturation logic
*)

(* CONTRACT_RULES [] *)

recipeAdded    := FALSE;
recipeDeleted  := FALSE;
recipeModified := FALSE;
local_opExecuted := FALSE;

IF queryRecipe THEN
    local_opExecuted := TRUE;
    error  := FALSE;
    status := 16#0000;
    local_found := FALSE;

    FOR local_index := 1 TO 10 DO
        IF recipe[local_index].recipeID = recipeIn.recipeID THEN
            local_found := TRUE;
            EXIT;
        END_IF;
    END_FOR;

    IF local_found THEN
        recipeQueryResult := recipe[local_index];
    ELSE
        error  := TRUE;
        status := 16#8001;
    END_IF;
END_IF;

IF addRecipe THEN
    local_opExecuted := TRUE;
    error  := FALSE;
    status := 16#0000;
    local_found    := FALSE;
    local_hasEmpty := FALSE;
    local_emptySlot := 0;

    FOR local_index := 1 TO 10 DO
        IF recipe[local_index].recipeID = recipeIn.recipeID THEN
            local_found := TRUE;
            EXIT;
        END_IF;
        IF recipe[local_index].recipeID = 0 AND NOT local_hasEmpty THEN
            local_hasEmpty  := TRUE;
            local_emptySlot := local_index;
        END_IF;
    END_FOR;

    IF local_found THEN
        error  := TRUE;
        status := 16#8002;
    ELSIF NOT local_hasEmpty THEN
        error  := TRUE;
        status := 16#8003;
    ELSE
        recipe[local_emptySlot] := recipeIn;
        recipeAdded             := TRUE;
    END_IF;
END_IF;

IF deleteRecipe THEN
    local_opExecuted := TRUE;
    error  := FALSE;
    status := 16#0000;
    local_found := FALSE;

    FOR local_index := 1 TO 10 DO
        IF recipe[local_index].recipeID = recipeIn.recipeID THEN
            local_found := TRUE;
            EXIT;
        END_IF;
    END_FOR;

    IF local_found THEN
        recipe[local_index].recipeID := 0;
        recipeDeleted                := TRUE;
    ELSE
        error  := TRUE;
        status := 16#8004;
    END_IF;
END_IF;

IF modifyRecipe THEN
    local_opExecuted := TRUE;
    error  := FALSE;
    status := 16#0000;
    local_found := FALSE;

    FOR local_index := 1 TO 10 DO
        IF recipe[local_index].recipeID = recipeIn.recipeID THEN
            local_found := TRUE;
            EXIT;
        END_IF;
    END_FOR;

    IF local_found THEN
        recipe[local_index] := recipeIn;
        recipeModified      := TRUE;
    ELSE
        error  := TRUE;
        status := 16#8005;
    END_IF;
END_IF;

END_FUNCTION_BLOCK

(* ---- public-hard-03.raw_candidate_01.st ---- *)
{+
Engineer: Claude
Date: 2026-11-13
Purpose: Recipe Management System per task specification
-}
FUNCTION_BLOCK FB_RecipeManager
VAR_INPUT
    addRecipe    : BOOL;
    deleteRecipe : BOOL;
    modifyRecipe : BOOL;
    queryRecipe  : BOOL;
    recipeIn     : ST_Recipe;
END_VAR
VAR_OUTPUT
    recipeAdded       : BOOL := FALSE;
    recipeDeleted     : BOOL := FALSE;
    recipeModified    : BOOL := FALSE;
    error             : BOOL := FALSE;
    status            : WORD := 16#0000;
    recipeQueryResult : ST_Recipe;
END_VAR
VAR_IN_OUT
    recipe : ARRAY[1..10] OF ST_Recipe;
END_VAR
VAR
    tmp_index     : INT;
    tmp_found     : BOOL;
    tmp_emptySlot : INT;
    tmp_hasEmpty  : BOOL;
END_VAR

(*
ENGINEERING_CONTRACT
====================
Operation Execution (same-scan, sequential priority order):
1. queryRecipe  → PUB001, PUB002, PUB008
2. addRecipe    → PUB002, PUB003, PUB009
3. deleteRecipe → PUB002, PUB004, PUB010
4. modifyRecipe → PUB002, PUB005, PUB011

Outputs - Activation/Retention/Reset:
- recipeAdded/recipeDeleted/recipeModified: pulse TRUE on success for current scan only (no retention)
- error: TRUE when any error occurs; no explicit reset (overwritten next scan)
- status: 16#0000 no-error, or error code 16#8001-16#8005 per PUB002

Error Codes (PUB002):
- 16#8001: queryRecipe - recipeID not found
- 16#8002: addRecipe   - recipeID already exists (duplicate)
- 16#8003: addRecipe   - no empty slot (database full)
- 16#8004: deleteRecipe - recipeID not found
- 16#8005: modifyRecipe - recipeID not found

Database Semantics (PUB006, PUB007):
- Array index range: [1..10], fixed
- Empty slot: recipeID = 0
- Add stores at smallest index empty slot (lowest array index)
- Delete sets recipeID to 0 (marks slot empty)
- Duplicate recipeID prohibited

Boundary Checks:
- recipeID comparisons use exact equality
- No wraparound or saturation logic
*)

(* CONTRACT_RULES [] *)

recipeAdded    := FALSE;
recipeDeleted  := FALSE;
recipeModified := FALSE;
error          := FALSE;
status         := 16#0000;

IF queryRecipe THEN
    tmp_found  := FALSE;
    tmp_index  := 1;
    FOR tmp_index := 1 TO 10 DO
        IF recipe[tmp_index].recipeID = recipeIn.recipeID THEN
            tmp_found := TRUE;
            EXIT;
        END_IF
    END_FOR;

    IF tmp_found THEN
        recipeQueryResult := recipe[tmp_index];
    ELSE
        error  := TRUE;
        status := 16#8001;
    END_IF;
END_IF;

IF addRecipe THEN
    tmp_found     := FALSE;
    tmp_hasEmpty  := FALSE;
    tmp_emptySlot := 0;

    FOR tmp_index := 1 TO 10 DO
        IF recipe[tmp_index].recipeID = recipeIn.recipeID THEN
            tmp_found := TRUE;
            EXIT;
        END_IF;
        IF recipe[tmp_index].recipeID = 0 AND NOT tmp_hasEmpty THEN
            tmp_hasEmpty  := TRUE;
            tmp_emptySlot := tmp_index;
        END_IF;
    END_FOR;

    IF tmp_found THEN
        error  := TRUE;
        status := 16#8002;
    ELSIF NOT tmp_hasEmpty THEN
        error  := TRUE;
        status := 16#8003;
    ELSE
        recipe[tmp_emptySlot] := recipeIn;
        recipeAdded           := TRUE;
    END_IF;
END_IF;

IF deleteRecipe THEN
    tmp_found := FALSE;
    tmp_index := 1;

    FOR tmp_index := 1 TO 10 DO
        IF recipe[tmp_index].recipeID = recipeIn.recipeID THEN
            tmp_found := TRUE;
            EXIT;
        END_IF;
    END_FOR;

    IF tmp_found THEN
        recipe[tmp_index].recipeID := 0;
        recipeDeleted              := TRUE;
    ELSE
        error  := TRUE;
        status := 16#8004;
    END_IF;
END_IF;

IF modifyRecipe THEN
    tmp_found := FALSE;
    tmp_index := 1;

    FOR tmp_index := 1 TO 10 DO
        IF recipe[tmp_index].recipeID = recipeIn.recipeID THEN
            tmp_found := TRUE;
            EXIT;
        END_IF;
    END_FOR;

    IF tmp_found THEN
        recipe[tmp_index] := recipeIn;
        recipeModified    := TRUE;
    ELSE
        error  := TRUE;
        status := 16#8005;
    END_IF;
END_IF;

END_FUNCTION_BLOCK

(* ---- public-hard-03.raw_candidate_02.st ---- *)
{+
FUNCTION_BLOCK FB_RecipeManager
VAR_INPUT
    addRecipe    : BOOL;
    deleteRecipe : BOOL;
    modifyRecipe : BOOL;
    queryRecipe  : BOOL;
    recipeIn     : ST_Recipe;
END_VAR
VAR_OUTPUT
    recipeAdded       : BOOL := FALSE;
    recipeDeleted     : BOOL := FALSE;
    recipeModified    : BOOL := FALSE;
    error             : BOOL := FALSE;
    status            : WORD := 16#0000;
    recipeQueryResult : ST_Recipe;
END_VAR
VAR_IN_OUT
    recipe : ARRAY[1..10] OF ST_Recipe;
END_VAR
VAR
    tmp_index     : INT;
    tmp_found     : BOOL;
    tmp_emptySlot : INT;
    tmp_hasEmpty  : BOOL;
END_VAR

(* ENGINEERING_CONTRACT
   ====================
   Operation Execution (same-scan, sequential priority):
   1. queryRecipe  → PUB008
   2. addRecipe    → PUB009
   3. deleteRecipe → PUB010
   4. modifyRecipe → PUB011

   Outputs - Activation/Retention/Reset:
   - recipeAdded/recipeDeleted/recipeModified: pulse TRUE on success for current scan only
   - error: TRUE when any error occurs; no explicit reset (overwritten next scan)
   - status: 16#0000 no-error, or error code 16#8001-16#8005 per PUB002

   Error Codes (PUB002):
   - 16#8001: queryRecipe - recipeID not found
   - 16#8002: addRecipe   - recipeID already exists (duplicate)
   - 16#8003: addRecipe   - no empty slot (database full)
   - 16#8004: deleteRecipe - recipeID not found
   - 16#8005: modifyRecipe - recipeID not found

   Database Semantics (PUB006, PUB007):
   - Array index range: [1..10], fixed
   - Empty slot: recipeID = 0
   - Add stores at smallest index empty slot
   - Delete sets recipeID to 0 (marks slot empty)
   - Duplicate recipeID prohibited
*)

(* CONTRACT_RULES [] *)

recipeAdded    := FALSE;
recipeDeleted  := FALSE;
recipeModified := FALSE;
error          := FALSE;
status         := 16#0000;

IF queryRecipe THEN
    tmp_found := FALSE;
    tmp_index := 1;
    WHILE tmp_index <= 10 AND NOT tmp_found DO
        IF recipe[tmp_index].recipeID = recipeIn.recipeID THEN
            tmp_found := TRUE;
        ELSE
            tmp_index := tmp_index + 1;
        END_IF;
    END_WHILE;

    IF tmp_found THEN
        recipeQueryResult := recipe[tmp_index];
    ELSE
        error  := TRUE;
        status := 16#8001;
    END_IF;
END_IF;

IF addRecipe THEN
    tmp_found     := FALSE;
    tmp_hasEmpty  := FALSE;
    tmp_emptySlot := 0;
    tmp_index     := 1;

    WHILE tmp_index <= 10 DO
        IF recipe[tmp_index].recipeID = recipeIn.recipeID THEN
            tmp_found := TRUE;
            tmp_index := 11;
        ELSE
            IF recipe[tmp_index].recipeID = 0 AND NOT tmp_hasEmpty THEN
                tmp_hasEmpty  := TRUE;
                tmp_emptySlot := tmp_index;
            END_IF;
            tmp_index := tmp_index + 1;
        END_IF;
    END_WHILE;

    IF tmp_found THEN
        error  := TRUE;
        status := 16#8002;
    ELSIF NOT tmp_hasEmpty THEN
        error  := TRUE;
        status := 16#8003;
    ELSE
        recipe[tmp_emptySlot] := recipeIn;
        recipeAdded           := TRUE;
    END_IF;
END_IF;

IF deleteRecipe THEN
    tmp_found := FALSE;
    tmp_index := 1;

    WHILE tmp_index <= 10 AND NOT tmp_found DO
        IF recipe[tmp_index].recipeID = recipeIn.recipeID THEN
            tmp_found := TRUE;
        ELSE
            tmp_index := tmp_index + 1;
        END_IF;
    END_WHILE;

    IF tmp_found THEN
        recipe[tmp_index].recipeID := 0;
        recipeDeleted              := TRUE;
    ELSE
        error  := TRUE;
        status := 16#8004;
    END_IF;
END_IF;

IF modifyRecipe THEN
    tmp_found := FALSE;
    tmp_index := 1;

    WHILE tmp_index <= 10 AND NOT tmp_found DO
        IF recipe[tmp_index].recipeID = recipeIn.recipeID THEN
            tmp_found := TRUE;
        ELSE
            tmp_index := tmp_index + 1;
        END_IF;
    END_WHILE;

    IF tmp_found THEN
        recipe[tmp_index] := recipeIn;
        recipeModified    := TRUE;
    ELSE
        error  := TRUE;
        status := 16#8005;
    END_IF;
END_IF;

END_FUNCTION_BLOCK
}

(* ---- public-hard-03.raw_candidate_03.st ---- *)
TYPE ST_Recipe :
STRUCT
    recipeID              : INT;
    ingredientType        : INT;
    ingredientRatio       : REAL;
    productionTemperature : REAL;
END_STRUCT
END_TYPE

FUNCTION_BLOCK FB_RecipeManager
VAR_INPUT
    addRecipe    : BOOL;
    deleteRecipe : BOOL;
    modifyRecipe : BOOL;
    queryRecipe  : BOOL;
    recipeIn     : ST_Recipe;
END_VAR
VAR_OUTPUT
    recipeAdded       : BOOL := FALSE;
    recipeDeleted     : BOOL := FALSE;
    recipeModified    : BOOL := FALSE;
    error             : BOOL := FALSE;
    status            : WORD := 16#0000;
    recipeQueryResult : ST_Recipe;
END_VAR
VAR_IN_OUT
    recipe : ARRAY[1..10] OF ST_Recipe;
END_VAR
VAR
    tmp_index     : INT;
    tmp_found     : BOOL;
    tmp_emptySlot : INT;
    tmp_hasEmpty  : BOOL;
END_VAR

(*
ENGINEERING_CONTRACT
====================
Operation Execution (same-scan, sequential priority order):
1. queryRecipe  -> PUB001, PUB002, PUB008
2. addRecipe    -> PUB002, PUB003, PUB009
3. deleteRecipe -> PUB002, PUB004, PUB010
4. modifyRecipe -> PUB002, PUB005, PUB011

Outputs - Activation/Retention/Reset:
- recipeAdded/recipeDeleted/recipeModified: pulse TRUE on success for current scan only (no retention)
- error: TRUE when any error occurs; no explicit reset (overwritten next scan)
- status: 16#0000 no-error, or error code 16#8001-16#8005 per PUB002

Error Codes (PUB002):
- 16#8001: queryRecipe - recipeID not found
- 16#8002: addRecipe   - recipeID already exists (duplicate)
- 16#8003: addRecipe   - no empty slot (database full)
- 16#8004: deleteRecipe - recipeID not found
- 16#8005: modifyRecipe - recipeID not found

Database Semantics (PUB006, PUB007):
- Array index range: [1..10], fixed
- Empty slot: recipeID = 0
- Add stores at smallest index empty slot (lowest array index)
- Delete sets recipeID to 0 (marks slot empty)
- Duplicate recipeID prohibited

Boundary Checks:
- recipeID comparisons use exact equality
- No wraparound or saturation logic
*)

(* CONTRACT_RULES [] *)

recipeAdded    := FALSE;
recipeDeleted  := FALSE;
recipeModified := FALSE;
error          := FALSE;
status         := 16#0000;

IF queryRecipe THEN
    tmp_found := FALSE;

    FOR tmp_index := 1 TO 10 DO
        IF recipe[tmp_index].recipeID = recipeIn.recipeID THEN
            tmp_found := TRUE;
            EXIT;
        END_IF
    END_FOR;

    IF tmp_found THEN
        recipeQueryResult := recipe[tmp_index];
    ELSE
        error  := TRUE;
        status := 16#8001;
    END_IF;
END_IF;

IF addRecipe THEN
    tmp_found     := FALSE;
    tmp_hasEmpty  := FALSE;
    tmp_emptySlot := 0;

    FOR tmp_index := 1 TO 10 DO
        IF recipe[tmp_index].recipeID = recipeIn.recipeID THEN
            tmp_found := TRUE;
            EXIT;
        END_IF;
        IF recipe[tmp_index].recipeID = 0 AND NOT tmp_hasEmpty THEN
            tmp_hasEmpty  := TRUE;
            tmp_emptySlot := tmp_index;
        END_IF;
    END_FOR;

    IF tmp_found THEN
        error  := TRUE;
        status := 16#8002;
    ELSIF NOT tmp_hasEmpty THEN
        error  := TRUE;
        status := 16#8003;
    ELSE
        recipe[tmp_emptySlot] := recipeIn;
        recipeAdded           := TRUE;
    END_IF;
END_IF;

IF deleteRecipe THEN
    tmp_found := FALSE;

    FOR tmp_index := 1 TO 10 DO
        IF recipe[tmp_index].recipeID = recipeIn.recipeID THEN
            tmp_found := TRUE;
            EXIT;
        END_IF;
    END_FOR;

    IF tmp_found THEN
        recipe[tmp_index].recipeID := 0;
        recipeDeleted              := TRUE;
    ELSE
        error  := TRUE;
        status := 16#8004;
    END_IF;
END_IF;

IF modifyRecipe THEN
    tmp_found := FALSE;

    FOR tmp_index := 1 TO 10 DO
        IF recipe[tmp_index].recipeID = recipeIn.recipeID THEN
            tmp_found := TRUE;
            EXIT;
        END_IF;
    END_FOR;

    IF tmp_found THEN
        recipe[tmp_index] := recipeIn;
        recipeModified    := TRUE;
    ELSE
        error  := TRUE;
        status := 16#8005;
    END_IF;
END_IF;

END_FUNCTION_BLOCK

(* ---- public-hard-03.raw_candidate_04.st ---- *)
TYPE ST_Recipe :
STRUCT
    recipeID              : INT;
    ingredientType        : INT;
    ingredientRatio       : REAL;
    productionTemperature : REAL;
END_STRUCT
END_TYPE

FUNCTION_BLOCK FB_RecipeManager
VAR_INPUT
    addRecipe    : BOOL;
    deleteRecipe : BOOL;
    modifyRecipe : BOOL;
    queryRecipe  : BOOL;
    recipeIn     : ST_Recipe;
END_VAR
VAR_OUTPUT
    recipeAdded       : BOOL := FALSE;
    recipeDeleted     : BOOL := FALSE;
    recipeModified    : BOOL := FALSE;
    error             : BOOL := FALSE;
    status            : WORD := 16#0000;
    recipeQueryResult : ST_Recipe;
END_VAR
VAR_IN_OUT
    recipe : ARRAY[1..10] OF ST_Recipe;
END_VAR
VAR
    local_index         : INT;
    local_found         : BOOL;
    local_emptySlot     : INT;
    local_hasEmpty      : BOOL;
    local_opExecuted    : BOOL;
END_VAR

(*
ENGINEERING_CONTRACT
====================
Operation Execution (same-scan, sequential priority order):
1. queryRecipe  -> PUB001, PUB002, PUB008
2. addRecipe    -> PUB002, PUB003, PUB009
3. deleteRecipe -> PUB002, PUB004, PUB010
4. modifyRecipe -> PUB002, PUB005, PUB011

Outputs - Activation/Retention/Reset:
- recipeAdded/recipeDeleted/recipeModified: pulse TRUE on success for current scan only (no retention)
- error: TRUE when any error occurs; retained across calls until next operation runs
- status: 16#0000 no-error, or error code 16#8001-16#8005 per PUB002; retained across calls

Error Codes (PUB002):
- 16#8001: queryRecipe  - recipeID not found
- 16#8002: addRecipe    - recipeID already exists (duplicate)
- 16#8003: addRecipe    - no empty slot (database full)
- 16#8004: deleteRecipe - recipeID not found
- 16#8005: modifyRecipe - recipeID not found

Database Semantics (PUB006, PUB007):
- Array index range: [1..10], fixed
- Empty slot: recipeID = 0
- Add stores at smallest index empty slot (lowest array index)
- Delete sets recipeID to 0 (marks slot empty)
- Duplicate recipeID prohibited

Boundary Checks:
- recipeID comparisons use exact equality
- No wraparound or saturation logic
*)

(* CONTRACT_RULES [] *)

recipeAdded    := FALSE;
recipeDeleted  := FALSE;
recipeModified := FALSE;
local_opExecuted := FALSE;

IF queryRecipe THEN
    local_opExecuted := TRUE;
    error  := FALSE;
    status := 16#0000;
    local_found := FALSE;

    FOR local_index := 1 TO 10 DO
        IF recipe[local_index].recipeID = recipeIn.recipeID THEN
            local_found := TRUE;
            EXIT;
        END_IF;
    END_FOR;

    IF local_found THEN
        recipeQueryResult := recipe[local_index];
    ELSE
        error  := TRUE;
        status := 16#8001;
    END_IF;
END_IF;

IF addRecipe THEN
    local_opExecuted := TRUE;
    error  := FALSE;
    status := 16#0000;
    local_found    := FALSE;
    local_hasEmpty := FALSE;
    local_emptySlot := 0;

    FOR local_index := 1 TO 10 DO
        IF recipe[local_index].recipeID = recipeIn.recipeID THEN
            local_found := TRUE;
            EXIT;
        END_IF;
        IF recipe[local_index].recipeID = 0 AND NOT local_hasEmpty THEN
            local_hasEmpty  := TRUE;
            local_emptySlot := local_index;
        END_IF;
    END_FOR;

    IF local_found THEN
        error  := TRUE;
        status := 16#8002;
    ELSIF NOT local_hasEmpty THEN
        error  := TRUE;
        status := 16#8003;
    ELSE
        recipe[local_emptySlot] := recipeIn;
        recipeAdded             := TRUE;
    END_IF;
END_IF;

IF deleteRecipe THEN
    local_opExecuted := TRUE;
    error  := FALSE;
    status := 16#0000;
    local_found := FALSE;

    FOR local_index := 1 TO 10 DO
        IF recipe[local_index].recipeID = recipeIn.recipeID THEN
            local_found := TRUE;
            EXIT;
        END_IF;
    END_FOR;

    IF local_found THEN
        recipe[local_index].recipeID := 0;
        recipeDeleted                := TRUE;
    ELSE
        error  := TRUE;
        status := 16#8004;
    END_IF;
END_IF;

IF modifyRecipe THEN
    local_opExecuted := TRUE;
    error  := FALSE;
    status := 16#0000;
    local_found := FALSE;

    FOR local_index := 1 TO 10 DO
        IF recipe[local_index].recipeID = recipeIn.recipeID THEN
            local_found := TRUE;
            EXIT;
        END_IF;
    END_FOR;

    IF local_found THEN
        recipe[local_index] := recipeIn;
        recipeModified      := TRUE;
    ELSE
        error  := TRUE;
        status := 16#8005;
    END_IF;
END_IF;

END_FUNCTION_BLOCK

(* ---- public-hard-04.candidate_01.st ---- *)
(* CONTRACT_RULES [] *)
FUNCTION_BLOCK FB_FIFOQueue
VAR_INPUT
    enqueue  : BOOL;
    dequeue  : BOOL;
    reset    : BOOL;
END_VAR
VAR_OUTPUT
    elementCount : DINT := 0;
    status       : WORD := 16#0000;
END_VAR
VAR_IN_OUT
    item   : VARIANT;
    buffer : VARIANT;
END_VAR
VAR
    local_head    : DINT  := 0;
    local_tail    : DINT  := 0;
    local_capacity : DINT  := 0;
    local_firstCycle : BOOL := TRUE;
    local_enqueueTrig : R_TRIG;
    local_dequeueTrig : R_TRIG;
END_VAR

// ENGINEERING_CONTRACT
// =============================================================================
// Activation: R_TRIG on enqueue/dequeue detect rising edges only.
// Retention:  local_head, local_tail, elementCount persist across scans.
// Reset:      Any scan where reset=TRUE empties queue regardless of other inputs.
// Same-scan:  Reset > Enqueue > Dequeue priority chain; only one operation per scan.
// Boundaries: Capacity derived from buffer array bounds; elementCount [0..capacity].
// Status:     16#0000 idle/success, 16#8001 empty-dequeue, 16#8002 full-enqueue.
// =============================================================================

// Rising-edge detection on command inputs
local_enqueueTrig(CLK := enqueue);
local_dequeueTrig(CLK := dequeue);

// First invocation: initialize capacity from buffer array bounds
IF local_firstCycle THEN
    local_firstCycle := FALSE;
    local_capacity := __GETUB(buffer, 0) - __GETLB(buffer, 0) + 1;
    local_head := 0;
    local_tail := 0;
    elementCount := 0;
    status := 16#0000;
    RETURN;
END_IF;

// Reset: priority over enqueue/dequeue
IF reset THEN
    local_head := 0;
    local_tail := 0;
    elementCount := 0;
    status := 16#0000;
    RETURN;
END_IF;

// Enqueue request: rising edge + not full
IF local_enqueueTrig.Q THEN
    IF elementCount < local_capacity THEN
        // Append item at tail position
        buffer[local_tail] := item;
        local_tail := (local_tail + 1) MOD local_capacity;
        elementCount := elementCount + 1;
        status := 16#0000;
    ELSE
        status := 16#8002; // Full rejection
    END_IF;
    RETURN;
END_IF;

// Dequeue request: rising edge + not empty
IF local_dequeueTrig.Q THEN
    IF elementCount > 0 THEN
        // Retrieve and remove front element
        item := buffer[local_head];
        local_head := (local_head + 1) MOD local_capacity;
        elementCount := elementCount - 1;
        status := 16#0000;
    ELSE
        status := 16#8001; // Empty rejection
    END_IF;
    RETURN;
END_IF;

// Idle scan: no pending operation
status := 16#0000;
END_FUNCTION_BLOCK

(* ---- public-hard-04.candidate_02.st ---- *)
(* CONTRACT_RULES [] *)
FUNCTION_BLOCK FB_FIFOQueue
VAR_INPUT
    enqueue  : BOOL;
    dequeue  : BOOL;
    reset    : BOOL;
END_VAR
VAR_OUTPUT
    elementCount : DINT := 0;
    status       : WORD := 16#0000;
END_VAR
VAR_IN_OUT
    item   : VARIANT;
    buffer : VARIANT;
END_VAR
VAR
    local_head         : DINT  := 0;
    local_tail         : DINT  := 0;
    local_capacity     : DINT  := 0;
    local_firstCycle   : BOOL  := TRUE;
    local_enqueueTrig  : R_TRIG;
    local_dequeueTrig  : R_TRIG;
END_VAR

// ENGINEERING_CONTRACT
// =============================================================================
// Activation: R_TRIG on enqueue/dequeue detect rising edges only.
// Retention:  local_head, local_tail, elementCount persist across scans.
// Reset:      Any scan where reset=TRUE empties queue regardless of other inputs.
// Same-scan:  Reset > Enqueue > Dequeue priority chain; only one operation per scan.
// Boundaries: Capacity derived from buffer array bounds; elementCount [0..capacity].
// Status:     16#0000 idle/success, 16#8001 empty-dequeue, 16#8002 full-enqueue.
// =============================================================================

// Rising-edge detection on command inputs
local_enqueueTrig(CLK := enqueue);
local_dequeueTrig(CLK := dequeue);

// First invocation: initialize capacity from buffer array bounds
IF local_firstCycle THEN
    local_firstCycle := FALSE;
    local_capacity := TO_DINT(UPPER_BOUND(buffer, 1) - LOWER_BOUND(buffer, 1) + 1);
    local_head := 0;
    local_tail := 0;
    elementCount := 0;
    status := 16#0000;
    RETURN;
END_IF;

// Reset: priority over enqueue/dequeue
IF reset THEN
    local_head := 0;
    local_tail := 0;
    elementCount := 0;
    status := 16#0000;
    RETURN;
END_IF;

// Enqueue request: rising edge + not full
IF local_enqueueTrig.Q THEN
    IF elementCount < local_capacity THEN
        // Append item at tail position
        buffer[local_tail] := item;
        local_tail := (local_tail + 1) MOD local_capacity;
        elementCount := elementCount + 1;
        status := 16#0000;
    ELSE
        status := 16#8002; // Full rejection
    END_IF;
    RETURN;
END_IF;

// Dequeue request: rising edge + not empty
IF local_dequeueTrig.Q THEN
    IF elementCount > 0 THEN
        // Retrieve and remove front element
        item := buffer[local_head];
        local_head := (local_head + 1) MOD local_capacity;
        elementCount := elementCount - 1;
        status := 16#0000;
    ELSE
        status := 16#8001; // Empty rejection
    END_IF;
    RETURN;
END_IF;

// Idle scan: no pending operation
status := 16#0000;
END_FUNCTION_BLOCK

(* ---- public-hard-04.candidate_03.st ---- *)
(* CONTRACT_RULES [] *)
FUNCTION_BLOCK FB_FIFOQueue
VAR_INPUT
    enqueue  : BOOL;
    dequeue  : BOOL;
    reset    : BOOL;
END_VAR
VAR_OUTPUT
    elementCount : DINT := 0;
    status       : WORD := 16#0000;
END_VAR
VAR_IN_OUT
    item   : VARIANT;
    buffer : VARIANT;
END_VAR
VAR
    local_head        : DINT  := 0;
    local_tail        : DINT  := 0;
    local_capacity    : DINT  := 0;
    local_firstCycle  : BOOL  := TRUE;
    local_enqueueTrig : R_TRIG;
    local_dequeueTrig : R_TRIG;
END_VAR

// ENGINEERING_CONTRACT
// =============================================================================
// PUB001: Capacity derived from buffer array length; element type from array.
// PUB002: Enqueue on rising edge, append if not full; tail advances circularly.
// PUB003: Dequeue on rising edge, retrieve front if not empty; head advances.
// PUB004: Reset clears queue; takes priority; buffer values need not be cleared.
// PUB005: elementCount [0..capacity] reports valid elements; zero = empty.
// PUB006: Status 16#0000 idle/success, 16#8001 empty-dequeue, 16#8002 full-enqueue.
// PUB007: Caller must not enqueue and dequeue same scan; no interlock enforced.
// PUB008: Queue empty on first invocation; firstCycle init on first call.
// PUB009-PUB011: Status codes as defined.
// Activation: R_TRIG on enqueue/dequeue; state persists across scans.
// Retention: head, tail, elementCount held; reset clears them.
// Reset priority: reset > enqueue > dequeue > idle; one operation per scan.
// Boundaries: Capacity from LOWER/UPPER_BOUND; indices MOD capacity.
// =============================================================================

// Rising-edge detection
local_enqueueTrig(CLK := enqueue);
local_dequeueTrig(CLK := dequeue);

// First invocation: derive capacity from buffer array bounds
IF local_firstCycle THEN
    local_firstCycle := FALSE;
    local_capacity := TO_DINT(UPPER_BOUND(buffer, 1) - LOWER_BOUND(buffer, 1) + 1);
    local_head := 0;
    local_tail := 0;
    elementCount := 0;
    status := 16#0000;
    RETURN;
END_IF;

// Reset: highest priority
IF reset THEN
    local_head := 0;
    local_tail := 0;
    elementCount := 0;
    status := 16#0000;
    RETURN;
END_IF;

// Enqueue request
IF local_enqueueTrig.Q THEN
    IF elementCount < local_capacity THEN
        buffer[local_tail] := item;
        local_tail := (local_tail + 1) MOD local_capacity;
        elementCount := elementCount + 1;
        status := 16#0000;
    ELSE
        status := 16#8002;
    END_IF;
    RETURN;
END_IF;

// Dequeue request
IF local_dequeueTrig.Q THEN
    IF elementCount > 0 THEN
        item := buffer[local_head];
        local_head := (local_head + 1) MOD local_capacity;
        elementCount := elementCount - 1;
        status := 16#0000;
    ELSE
        status := 16#8001;
    END_IF;
    RETURN;
END_IF;

// Idle scan
status := 16#0000;
END_FUNCTION_BLOCK

(* ---- public-hard-04.candidate_04.st ---- *)
(* CONTRACT_RULES [] *)
FUNCTION_BLOCK FB_FIFOQueue
VAR_INPUT
    enqueue  : BOOL;
    dequeue  : BOOL;
    reset    : BOOL;
END_VAR
VAR_OUTPUT
    elementCount : DINT := 0;
    status       : WORD := 16#0000;
END_VAR
VAR_IN_OUT
    item   : VARIANT;
    buffer : VARIANT;
END_VAR
VAR
    local_head         : DINT  := 0;
    local_tail         : DINT  := 0;
    local_capacity     : DINT  := 0;
    local_firstCycle   : BOOL  := TRUE;
    local_enqueueTrig  : R_TRIG;
    local_dequeueTrig  : R_TRIG;
END_VAR

// ENGINEERING_CONTRACT
// =============================================================================
// Activation: R_TRIG on enqueue/dequeue detect rising edges only.
// Retention:  local_head, local_tail, elementCount persist across scans.
// Reset:      Any scan where reset=TRUE empties queue regardless of other inputs.
// Same-scan:  Reset > Enqueue > Dequeue priority chain; only one operation per scan.
// Boundaries: Capacity derived from buffer array bounds; elementCount [0..capacity].
// Status:     16#0000 idle/success, 16#8001 empty-dequeue, 16#8002 full-enqueue.
// =============================================================================

local_enqueueTrig(CLK := enqueue);
local_dequeueTrig(CLK := dequeue);

IF local_firstCycle THEN
    local_firstCycle := FALSE;
    local_capacity := TO_DINT(UPPER_BOUND(buffer, 1)) - TO_DINT(LOWER_BOUND(buffer, 1)) + 1;
    IF local_capacity <= 0 THEN
        local_capacity := 1;
    END_IF;
    local_head := 0;
    local_tail := 0;
    elementCount := 0;
    status := 16#0000;
    RETURN;
END_IF;

IF reset THEN
    local_head := 0;
    local_tail := 0;
    elementCount := 0;
    status := 16#0000;
    RETURN;
END_IF;

IF local_enqueueTrig.Q THEN
    IF elementCount < local_capacity THEN
        buffer[local_tail] := item;
        local_tail := (local_tail + 1) MOD local_capacity;
        elementCount := elementCount + 1;
        status := 16#0000;
    ELSE
        status := 16#8002;
    END_IF;
    RETURN;
END_IF;

IF local_dequeueTrig.Q THEN
    IF elementCount > 0 THEN
        item := buffer[local_head];
        local_head := (local_head + 1) MOD local_capacity;
        elementCount := elementCount - 1;
        status := 16#0000;
    ELSE
        status := 16#8001;
    END_IF;
    RETURN;
END_IF;

status := 16#0000;
END_FUNCTION_BLOCK

(* ---- public-hard-04.raw_candidate_01.st ---- *)
(* CONTRACT_RULES [] *)
FUNCTION_BLOCK FB_FIFOQueue
VAR_INPUT
    enqueue  : BOOL;
    dequeue  : BOOL;
    reset    : BOOL;
END_VAR
VAR_OUTPUT
    elementCount : DINT := 0;
    status       : WORD := 16#0000;
END_VAR
VAR_IN_OUT
    item   : VARIANT;
    buffer : VARIANT;
END_VAR
VAR
    local_head    : DINT  := 0;
    local_tail    : DINT  := 0;
    local_capacity : DINT  := 0;
    local_firstCycle : BOOL := TRUE;
    local_enqueueTrig : R_TRIG;
    local_dequeueTrig : R_TRIG;
END_VAR

// ENGINEERING_CONTRACT
// =============================================================================
// Activation: R_TRIG on enqueue/dequeue detect rising edges only.
// Retention:  local_head, local_tail, elementCount persist across scans.
// Reset:      Any scan where reset=TRUE empties queue regardless of other inputs.
// Same-scan:  Reset > Enqueue > Dequeue priority chain; only one operation per scan.
// Boundaries: Capacity derived from buffer array bounds; elementCount [0..capacity].
// Status:     16#0000 idle/success, 16#8001 empty-dequeue, 16#8002 full-enqueue.
// =============================================================================

// Rising-edge detection on command inputs
local_enqueueTrig(CLK := enqueue);
local_dequeueTrig(CLK := dequeue);

// First invocation: initialize capacity from buffer array bounds
IF local_firstCycle THEN
    local_firstCycle := FALSE;
    local_capacity := __GETUB(buffer, 0) - __GETLB(buffer, 0) + 1;
    local_head := 0;
    local_tail := 0;
    elementCount := 0;
    status := 16#0000;
    RETURN;
END_IF;

// Reset: priority over enqueue/dequeue
IF reset THEN
    local_head := 0;
    local_tail := 0;
    elementCount := 0;
    status := 16#0000;
    RETURN;
END_IF;

// Enqueue request: rising edge + not full
IF local_enqueueTrig.Q THEN
    IF elementCount < local_capacity THEN
        // Append item at tail position
        buffer[local_tail] := item;
        local_tail := (local_tail + 1) MOD local_capacity;
        elementCount := elementCount + 1;
        status := 16#0000;
    ELSE
        status := 16#8002; // Full rejection
    END_IF;
    RETURN;
END_IF;

// Dequeue request: rising edge + not empty
IF local_dequeueTrig.Q THEN
    IF elementCount > 0 THEN
        // Retrieve and remove front element
        item := buffer[local_head];
        local_head := (local_head + 1) MOD local_capacity;
        elementCount := elementCount - 1;
        status := 16#0000;
    ELSE
        status := 16#8001; // Empty rejection
    END_IF;
    RETURN;
END_IF;

// Idle scan: no pending operation
status := 16#0000;
END_FUNCTION_BLOCK

(* ---- public-hard-04.raw_candidate_02.st ---- *)
(* CONTRACT_RULES [] *)
FUNCTION_BLOCK FB_FIFOQueue
VAR_INPUT
    enqueue  : BOOL;
    dequeue  : BOOL;
    reset    : BOOL;
END_VAR
VAR_OUTPUT
    elementCount : DINT := 0;
    status       : WORD := 16#0000;
END_VAR
VAR_IN_OUT
    item   : VARIANT;
    buffer : VARIANT;
END_VAR
VAR
    local_head         : DINT  := 0;
    local_tail         : DINT  := 0;
    local_capacity     : DINT  := 0;
    local_firstCycle   : BOOL  := TRUE;
    local_enqueueTrig  : R_TRIG;
    local_dequeueTrig  : R_TRIG;
END_VAR

// ENGINEERING_CONTRACT
// =============================================================================
// Activation: R_TRIG on enqueue/dequeue detect rising edges only.
// Retention:  local_head, local_tail, elementCount persist across scans.
// Reset:      Any scan where reset=TRUE empties queue regardless of other inputs.
// Same-scan:  Reset > Enqueue > Dequeue priority chain; only one operation per scan.
// Boundaries: Capacity derived from buffer array bounds; elementCount [0..capacity].
// Status:     16#0000 idle/success, 16#8001 empty-dequeue, 16#8002 full-enqueue.
// =============================================================================

// Rising-edge detection on command inputs
local_enqueueTrig(CLK := enqueue);
local_dequeueTrig(CLK := dequeue);

// First invocation: initialize capacity from buffer array bounds
IF local_firstCycle THEN
    local_firstCycle := FALSE;
    local_capacity := TO_DINT(UPPER_BOUND(buffer, 1) - LOWER_BOUND(buffer, 1) + 1);
    local_head := 0;
    local_tail := 0;
    elementCount := 0;
    status := 16#0000;
    RETURN;
END_IF;

// Reset: priority over enqueue/dequeue
IF reset THEN
    local_head := 0;
    local_tail := 0;
    elementCount := 0;
    status := 16#0000;
    RETURN;
END_IF;

// Enqueue request: rising edge + not full
IF local_enqueueTrig.Q THEN
    IF elementCount < local_capacity THEN
        // Append item at tail position
        buffer[local_tail] := item;
        local_tail := (local_tail + 1) MOD local_capacity;
        elementCount := elementCount + 1;
        status := 16#0000;
    ELSE
        status := 16#8002; // Full rejection
    END_IF;
    RETURN;
END_IF;

// Dequeue request: rising edge + not empty
IF local_dequeueTrig.Q THEN
    IF elementCount > 0 THEN
        // Retrieve and remove front element
        item := buffer[local_head];
        local_head := (local_head + 1) MOD local_capacity;
        elementCount := elementCount - 1;
        status := 16#0000;
    ELSE
        status := 16#8001; // Empty rejection
    END_IF;
    RETURN;
END_IF;

// Idle scan: no pending operation
status := 16#0000;
END_FUNCTION_BLOCK

(* ---- public-hard-04.raw_candidate_03.st ---- *)
(* CONTRACT_RULES [] *)
FUNCTION_BLOCK FB_FIFOQueue
VAR_INPUT
    enqueue  : BOOL;
    dequeue  : BOOL;
    reset    : BOOL;
END_VAR
VAR_OUTPUT
    elementCount : DINT := 0;
    status       : WORD := 16#0000;
END_VAR
VAR_IN_OUT
    item   : VARIANT;
    buffer : VARIANT;
END_VAR
VAR
    local_head        : DINT  := 0;
    local_tail        : DINT  := 0;
    local_capacity    : DINT  := 0;
    local_firstCycle  : BOOL  := TRUE;
    local_enqueueTrig : R_TRIG;
    local_dequeueTrig : R_TRIG;
END_VAR

// ENGINEERING_CONTRACT
// =============================================================================
// PUB001: Capacity derived from buffer array length; element type from array.
// PUB002: Enqueue on rising edge, append if not full; tail advances circularly.
// PUB003: Dequeue on rising edge, retrieve front if not empty; head advances.
// PUB004: Reset clears queue; takes priority; buffer values need not be cleared.
// PUB005: elementCount [0..capacity] reports valid elements; zero = empty.
// PUB006: Status 16#0000 idle/success, 16#8001 empty-dequeue, 16#8002 full-enqueue.
// PUB007: Caller must not enqueue and dequeue same scan; no interlock enforced.
// PUB008: Queue empty on first invocation; firstCycle init on first call.
// PUB009-PUB011: Status codes as defined.
// Activation: R_TRIG on enqueue/dequeue; state persists across scans.
// Retention: head, tail, elementCount held; reset clears them.
// Reset priority: reset > enqueue > dequeue > idle; one operation per scan.
// Boundaries: Capacity from LOWER/UPPER_BOUND; indices MOD capacity.
// =============================================================================

// Rising-edge detection
local_enqueueTrig(CLK := enqueue);
local_dequeueTrig(CLK := dequeue);

// First invocation: derive capacity from buffer array bounds
IF local_firstCycle THEN
    local_firstCycle := FALSE;
    local_capacity := TO_DINT(UPPER_BOUND(buffer, 1) - LOWER_BOUND(buffer, 1) + 1);
    local_head := 0;
    local_tail := 0;
    elementCount := 0;
    status := 16#0000;
    RETURN;
END_IF;

// Reset: highest priority
IF reset THEN
    local_head := 0;
    local_tail := 0;
    elementCount := 0;
    status := 16#0000;
    RETURN;
END_IF;

// Enqueue request
IF local_enqueueTrig.Q THEN
    IF elementCount < local_capacity THEN
        buffer[local_tail] := item;
        local_tail := (local_tail + 1) MOD local_capacity;
        elementCount := elementCount + 1;
        status := 16#0000;
    ELSE
        status := 16#8002;
    END_IF;
    RETURN;
END_IF;

// Dequeue request
IF local_dequeueTrig.Q THEN
    IF elementCount > 0 THEN
        item := buffer[local_head];
        local_head := (local_head + 1) MOD local_capacity;
        elementCount := elementCount - 1;
        status := 16#0000;
    ELSE
        status := 16#8001;
    END_IF;
    RETURN;
END_IF;

// Idle scan
status := 16#0000;
END_FUNCTION_BLOCK

(* ---- public-hard-04.raw_candidate_04.st ---- *)
(* CONTRACT_RULES [] *)
FUNCTION_BLOCK FB_FIFOQueue
VAR_INPUT
    enqueue  : BOOL;
    dequeue  : BOOL;
    reset    : BOOL;
END_VAR
VAR_OUTPUT
    elementCount : DINT := 0;
    status       : WORD := 16#0000;
END_VAR
VAR_IN_OUT
    item   : VARIANT;
    buffer : VARIANT;
END_VAR
VAR
    local_head         : DINT  := 0;
    local_tail         : DINT  := 0;
    local_capacity     : DINT  := 0;
    local_firstCycle   : BOOL  := TRUE;
    local_enqueueTrig  : R_TRIG;
    local_dequeueTrig  : R_TRIG;
END_VAR

// ENGINEERING_CONTRACT
// =============================================================================
// Activation: R_TRIG on enqueue/dequeue detect rising edges only.
// Retention:  local_head, local_tail, elementCount persist across scans.
// Reset:      Any scan where reset=TRUE empties queue regardless of other inputs.
// Same-scan:  Reset > Enqueue > Dequeue priority chain; only one operation per scan.
// Boundaries: Capacity derived from buffer array bounds; elementCount [0..capacity].
// Status:     16#0000 idle/success, 16#8001 empty-dequeue, 16#8002 full-enqueue.
// =============================================================================

local_enqueueTrig(CLK := enqueue);
local_dequeueTrig(CLK := dequeue);

IF local_firstCycle THEN
    local_firstCycle := FALSE;
    local_capacity := TO_DINT(UPPER_BOUND(buffer, 1)) - TO_DINT(LOWER_BOUND(buffer, 1)) + 1;
    IF local_capacity <= 0 THEN
        local_capacity := 1;
    END_IF;
    local_head := 0;
    local_tail := 0;
    elementCount := 0;
    status := 16#0000;
    RETURN;
END_IF;

IF reset THEN
    local_head := 0;
    local_tail := 0;
    elementCount := 0;
    status := 16#0000;
    RETURN;
END_IF;

IF local_enqueueTrig.Q THEN
    IF elementCount < local_capacity THEN
        buffer[local_tail] := item;
        local_tail := (local_tail + 1) MOD local_capacity;
        elementCount := elementCount + 1;
        status := 16#0000;
    ELSE
        status := 16#8002;
    END_IF;
    RETURN;
END_IF;

IF local_dequeueTrig.Q THEN
    IF elementCount > 0 THEN
        item := buffer[local_head];
        local_head := (local_head + 1) MOD local_capacity;
        elementCount := elementCount - 1;
        status := 16#0000;
    ELSE
        status := 16#8001;
    END_IF;
    RETURN;
END_IF;

status := 16#0000;
END_FUNCTION_BLOCK

(* ---- public-hard-05.candidate_01.st ---- *)
FUNCTION_BLOCK ArmController
VAR_INPUT
    ManualMode : BOOL;
    SingleStepMode : BOOL;
    SingleCycleMode : BOOL;
    ContinuousMode : BOOL;
    EmergencyStop : BOOL;
    Start : BOOL;
    DownButton : BOOL;
    UpButton : BOOL;
    LeftButton : BOOL;
    RightButton : BOOL;
    GripButton : BOOL;
    ReleaseButton : BOOL;
    DownLimitSwitch : BOOL;
    UpLimitSwitch : BOOL;
    LeftLimitSwitch : BOOL;
    RightLimitSwitch : BOOL;
    GripLimitSwitch : BOOL;
    ReleaseLimitSwitch : BOOL;
END_VAR
VAR_OUTPUT
    MoveDown : BOOL := FALSE;
    MoveUp : BOOL := FALSE;
    MoveLeft : BOOL := FALSE;
    MoveRight : BOOL := FALSE;
    ActivateGrip : BOOL := FALSE;
    ActivateRelease : BOOL := FALSE;
END_VAR
VAR
    step : INT := 0;
    startRisingEdge : R_TRIG;
    running : BOOL := FALSE;
    cycleComplete : BOOL := FALSE;
    tmpRunning : BOOL;
END_VAR

(* ENGINEERING_CONTRACT
| Output/State      | Activation       | Retention       | Reset/Deactivation             | Same-Scan Priority    | Units/Boundaries      |
|-------------------|------------------|-----------------|---------------------------------|-----------------------|-----------------------|
| MoveDown/Up/Left/Right | Edge/start/trig | Hold until done | EmergencyStop(FALSE), mode end  | Output latches stop   | BOOL, limit-based     |
| ActivateGrip/Release   | Edge/start/trig | Hold until done | EmergencyStop(FALSE), mode end  | Output latches stop   | BOOL, limit-based     |
| step[0..8]        | Start rising edge| Retained        | EmergencyStop(FALSE), mode end  | Initialized to 0      | INT, wrap to 0 at 8   |
| running           | Start rising edge| Retained        | EmergencyStop(FALSE), cycle end | FALSE when E-Stop     | BOOL, auto in cycle   |
| cycleComplete     | step=8 & done    | Retained        | Start rising edge               | Set only once         | BOOL, latched         |

PUB clause coverage:
- PUB001: Manual mode direct button control with limit checking
- PUB002-PUB007: Single step sequence (8 steps, Start advances)
- PUB008-PUB011: Single cycle executes full sequence once
- PUB012-PUB015: Continuous mode repeats cycle
- PUB016-PUB018: Emergency stop (FALSE=triggered) stops all outputs
- PUB019-PUB020: Grip/Release limit switches for completion feedback

Behavior:
- EmergencyStop=FALSE: All outputs=0, running=FALSE, step NOT reset (resume capability)
- Initial state: step=0, running=FALSE, all outputs=FALSE
- Caller ensures mutually exclusive mode inputs
*)
(* CONTRACT_RULES [] *)

tmpRunning := running;

startRisingEdge(CLK := Start);
running := running OR (startRisingEdge.Q AND (SingleStepMode OR SingleCycleMode OR ContinuousMode));

IF EmergencyStop = FALSE THEN
    MoveDown := FALSE;
    MoveUp := FALSE;
    MoveLeft := FALSE;
    MoveRight := FALSE;
    ActivateGrip := FALSE;
    ActivateRelease := FALSE;
    running := FALSE;
    cycleComplete := FALSE;
ELSE
    IF ManualMode THEN
        step := 0;
        running := FALSE;

        IF DownButton AND NOT DownLimitSwitch THEN
            MoveDown := TRUE;
        END_IF;
        IF UpButton AND NOT UpLimitSwitch THEN
            MoveUp := TRUE;
        END_IF;
        IF LeftButton AND NOT LeftLimitSwitch THEN
            MoveLeft := TRUE;
        END_IF;
        IF RightButton AND NOT RightLimitSwitch THEN
            MoveRight := TRUE;
        END_IF;
        IF GripButton THEN
            ActivateGrip := TRUE;
        END_IF;
        IF ReleaseButton THEN
            ActivateRelease := TRUE;
        END_IF;

    ELSIF SingleStepMode THEN
        IF startRisingEdge.Q AND NOT running THEN
            running := TRUE;
        END_IF;

        IF running THEN
            CASE step OF
                0:
                    IF UpLimitSwitch THEN
                        MoveDown := TRUE;
                        IF DownLimitSwitch THEN
                            MoveDown := FALSE;
                            step := 1;
                        END_IF;
                    END_IF;
                1:
                    MoveDown := FALSE;
                    ActivateGrip := TRUE;
                    IF GripLimitSwitch THEN
                        ActivateGrip := FALSE;
                        step := 2;
                    END_IF;
                2:
                    ActivateGrip := FALSE;
                    MoveUp := TRUE;
                    IF UpLimitSwitch THEN
                        MoveUp := FALSE;
                        step := 3;
                    END_IF;
                3:
                    MoveUp := FALSE;
                    MoveRight := TRUE;
                    IF RightLimitSwitch THEN
                        MoveRight := FALSE;
                        step := 4;
                    END_IF;
                4:
                    MoveRight := FALSE;
                    MoveDown := TRUE;
                    IF DownLimitSwitch THEN
                        MoveDown := FALSE;
                        step := 5;
                    END_IF;
                5:
                    MoveDown := FALSE;
                    ActivateRelease := TRUE;
                    IF ReleaseLimitSwitch THEN
                        ActivateRelease := FALSE;
                        step := 6;
                    END_IF;
                6:
                    ActivateRelease := FALSE;
                    MoveUp := TRUE;
                    IF UpLimitSwitch THEN
                        MoveUp := FALSE;
                        step := 7;
                    END_IF;
                7:
                    MoveUp := FALSE;
                    MoveLeft := TRUE;
                    IF LeftLimitSwitch THEN
                        MoveLeft := FALSE;
                        step := 8;
                    END_IF;
                8:
                    MoveLeft := FALSE;
                    running := FALSE;
                    step := 0;
            END_CASE;
        END_IF;

    ELSIF SingleCycleMode THEN
        IF startRisingEdge.Q AND NOT running AND NOT cycleComplete THEN
            running := TRUE;
        END_IF;

        IF running AND NOT cycleComplete THEN
            CASE step OF
                0:
                    IF UpLimitSwitch THEN
                        MoveDown := TRUE;
                        IF DownLimitSwitch THEN
                            MoveDown := FALSE;
                            step := 1;
                        END_IF;
                    END_IF;
                1:
                    MoveDown := FALSE;
                    ActivateGrip := TRUE;
                    IF GripLimitSwitch THEN
                        ActivateGrip := FALSE;
                        step := 2;
                    END_IF;
                2:
                    ActivateGrip := FALSE;
                    MoveUp := TRUE;
                    IF UpLimitSwitch THEN
                        MoveUp := FALSE;
                        step := 3;
                    END_IF;
                3:
                    MoveUp := FALSE;
                    MoveRight := TRUE;
                    IF RightLimitSwitch THEN
                        MoveRight := FALSE;
                        step := 4;
                    END_IF;
                4:
                    MoveRight := FALSE;
                    MoveDown := TRUE;
                    IF DownLimitSwitch THEN
                        MoveDown := FALSE;
                        step := 5;
                    END_IF;
                5:
                    MoveDown := FALSE;
                    ActivateRelease := TRUE;
                    IF ReleaseLimitSwitch THEN
                        ActivateRelease := FALSE;
                        step := 6;
                    END_IF;
                6:
                    ActivateRelease := FALSE;
                    MoveUp := TRUE;
                    IF UpLimitSwitch THEN
                        MoveUp := FALSE;
                        step := 7;
                    END_IF;
                7:
                    MoveUp := FALSE;
                    MoveLeft := TRUE;
                    IF LeftLimitSwitch THEN
                        MoveLeft := FALSE;
                        step := 8;
                    END_IF;
                8:
                    MoveLeft := FALSE;
                    running := FALSE;
                    cycleComplete := TRUE;
                    step := 0;
            END_CASE;
        END_IF;

    ELSIF ContinuousMode THEN
        IF startRisingEdge.Q AND NOT running THEN
            running := TRUE;
        END_IF;

        IF running THEN
            CASE step OF
                0:
                    IF UpLimitSwitch THEN
                        MoveDown := TRUE;
                        IF DownLimitSwitch THEN
                            MoveDown := FALSE;
                            step := 1;
                        END_IF;
                    END_IF;
                1:
                    MoveDown := FALSE;
                    ActivateGrip := TRUE;
                    IF GripLimitSwitch THEN
                        ActivateGrip := FALSE;
                        step := 2;
                    END_IF;
                2:
                    ActivateGrip := FALSE;
                    MoveUp := TRUE;
                    IF UpLimitSwitch THEN
                        MoveUp := FALSE;
                        step := 3;
                    END_IF;
                3:
                    MoveUp := FALSE;
                    MoveRight := TRUE;
                    IF RightLimitSwitch THEN
                        MoveRight := FALSE;
                        step := 4;
                    END_IF;
                4:
                    MoveRight := FALSE;
                    MoveDown := TRUE;
                    IF DownLimitSwitch THEN
                        MoveDown := FALSE;
                        step := 5;
                    END_IF;
                5:
                    MoveDown := FALSE;
                    ActivateRelease := TRUE;
                    IF ReleaseLimitSwitch THEN
                        ActivateRelease := FALSE;
                        step := 6;
                    END_IF;
                6:
                    ActivateRelease := FALSE;
                    MoveUp := TRUE;
                    IF UpLimitSwitch THEN
                        MoveUp := FALSE;
                        step := 7;
                    END_IF;
                7:
                    MoveUp := FALSE;
                    MoveLeft := TRUE;
                    IF LeftLimitSwitch THEN
                        MoveLeft := FALSE;
                        step := 0;
                    END_IF;
            END_CASE;
        END_IF;
    END_IF;
END_IF;

END_FUNCTION_BLOCK
